Fanuc KAREL source: KT00107.KL

PROGRAM KT00107
%NOLOCKGROUP
VAR
  R1: REAL
  R2: REAL
  OUT: INTEGER
BEGIN
  R1 = 2.0
  R2 = 3.0
  R1 = 2.0
  R2 = 3.0
  OUT = R1 / R2
END KT00107
